# EPICS substitutions: db/Beckhoff_7XXX/ecmcEL7211-0010_CSP.substitutions
file "ecmcEL72XX_DRV_CSP.template"
{
  pattern {CH_ID}
          {01   }
}

file "ecmcEL72XX_ENC.template"
{
  pattern {CH_ID}
          {01   }
}
